Fanuc KAREL source: kt00601.KL

-- PROVISIONAL review KL for V940-1; original PC SHA256 ad41c04657136a2a10db56503cc8705a3705e376cdb1fa6fac56468a867cf11e
-- Incomplete behavior may be omitted. Consult companion uncertainty JSON. Do not deploy.
PROGRAM KT00601
%NOLOCKGROUP
VAR
  I1 : INTEGER
  I2 : INTEGER
  OUT : INTEGER
BEGIN
  -- V9_ZERO_TABLE_METADATA_HINT layout=0001; no indexed target words; source/name/runtime held
  -- UNRESOLVED_PC offsets 5-16; opcodes 2E,23
  -- UNRESOLVED_PC offsets 21-32; opcodes 2E,23
  -- UNRESOLVED_PC offsets 37-48; opcodes 2E,23
  -- UNRESOLVED_PC offsets 53-64; opcodes 2E,23
  -- UNRESOLVED_PC offsets 69-81; opcodes 21,23
  -- UNRESOLVED_PC offsets 86-90; opcodes 7F
END KT00601
